{attribute 'qualified_only'}
VAR_GLOBAL
	
	// Lamp varibol
	OXLampOXOne :BOOL;
	OXLampIXOneGreen :BOOL;
	OXLampOXTwo :BOOL;
	OXLampIXTwoGreen :BOOL;
	
	//strob out
	oxStrobOne AT %Q* : BOOL ;
	oxStrobTwo AT %Q* : BOOL ;
 	//strob in
	ixStrobOne AT %I* : BOOL ;
	ixStrobTwo AT %I* : BOOL ;
	
	// Long or Short
	ixLong AT %I* : BOOL;
	ixShort AT%I* :BOOL;
	
	// car move
	OIntRedCar: INT;
	OintCopCar: INT;
END_VAR

(* stored: Version 1.1.0.1, ProductVersion 3.1.4024.12
   GVL GVLSlave: Id {840cc7fc-3cf5-4a40-8947-ce7af77b5757} *)
